{attribute 'qualified_only'}
VAR_GLOBAL
	Target_A : ARRAY [1..3] OF LREAL := [0.0, 200.0, 0.0];
    Target_B : ARRAY [1..3] OF LREAL := [450.0, 100.0, 30.0];
    Target_C : ARRAY [1..3] OF LREAL := [450.0, -100.0, -30.0];
END_VAR

(* stored: Version 1.1.0.1, ProductVersion 3.1.4024.15
   GVL GVL_TargetPoints: Id {0f09f3b1-3b1f-44c1-885b-7a5aae76a14e} *)
